// TIA Portal V20 export
// export: Created 2026-10-19T18:44:59.9625904Z, ExportSetting None, DisplayName Totally Integrated Automation Portal, DisplayVersion V20 Update 6, DisplayName TIA Portal Openness, DisplayVersion V20 Update 6, DisplayName TIA Portal Version Control Interface, DisplayVersion V20 Update 6, DisplayName SINAMICS Startdrive Advanced, DisplayVersion V20 SP1, DisplayName SINAMICS Startdrive G130, G150, S120, S150, SINAMICS MV, G220, S200, S210, DisplayVersion V20 SP1, DisplayName SINAMICS Startdrive G110M, G120, G120C, G120D, G120P, G115D, DisplayVersion V20 SP1, DisplayName STEP 7 Professional, DisplayVersion V20 Update 6, DisplayName STEP 7 Safety, DisplayVersion V20 Update 2, DisplayName WinCC Basic/Comfort/Advanced, DisplayVersion V20 Update 6, DisplayName WinCC Unified, DisplayVersion V20 Update 6
VAR_GLOBAL   // PLC tag table "Default tag table"
   System_Byte AT %MB1159 : Byte;
   FirstScan AT %M1159.0 : Bool;
   DiagStatusUpdate AT %M1159.1 : Bool;
   AlwaysTRUE AT %M1159.2 : Bool;
   AlwaysFALSE AT %M1159.3 : Bool;
   Clock_Byte AT %MB1160 : Byte;
   Clock_10Hz AT %M1160.0 : Bool;
   Clock_5Hz AT %M1160.1 : Bool;
   "Clock_2.5Hz" AT %M1160.2 : Bool;
   Clock_2Hz AT %M1160.3 : Bool;
   "Clock_1.25Hz" AT %M1160.4 : Bool;
   Clock_1Hz AT %M1160.5 : Bool;
   "Clock_0.625Hz" AT %M1160.6 : Bool;
   "Clock_0.5Hz" AT %M1160.7 : Bool;
   Tag_1 AT %M2000.0 : Bool;
   Tag_2 AT %M2000.1 : Bool;
   Tag_3 AT %M2000.2 : Bool;
   Reintegration AT %M2000.3 : Bool;
   Error_Word_1 AT %MW2001 : Word;
   "Auto_Stop_Lector(1)" AT %M20.6 : Bool;
   "Auto_Stop_Lector(2)" AT %M20.7 : Bool;
   "Auto_Start_Lector(1)" AT %M19.6 : Bool;
   "Auto_Start_Lector(2)" AT %M20.2 : Bool;
   Force_System_1 AT %M25.5 : Bool;
   VTD_System_Selected_HMI AT %MW1234 : UInt;
   Initialization AT %M19.4 : Bool;
   Save_Settings AT %M0.1 : Bool;
   "LE_Bypass(1)" AT %M704.1 : Bool;
   "LE_Bypass(2)" AT %M704.2 : Bool;
   Reset_Comissioning AT %M70.0 : Bool;
   System_2_Busy AT %M39.6 : Bool;
   System_1_Busy AT %M19.5 : Bool;
   L3_OK AT %M39.4 : Bool;
   L4_OK AT %M39.0 : Bool;
   L5_OK AT %M39.1 : Bool;
   L1_OK AT %M26.6 : Bool;
   L2_OK AT %M26.7 : Bool;
   L6_OK AT %M39.2 : Bool;
   L1_Estop AT %M61.6 : Bool;
   L6_Estop AT %M70.6 : Bool;
   L2_Estop AT %M61.7 : Bool;
   L5_Estop AT %M70.4 : Bool;
   L4_Estop AT %M70.3 : Bool;
   L3_Estop AT %M70.2 : Bool;
   LGX_Secure_Access_2 AT %M71.5 : Bool;
   LGX_Secure_Access_1 AT %M71.4 : Bool;
   LGX_ReadyToReceive_2 AT %M71.2 : Bool;
   LGX_ReadyToReceive_1 AT %M61.5 : Bool;
   Dbug AT %M71.7 : Bool;
   OrderNo AT %MW158 : Int;
   "Clear_OT_Buffers(1)" AT %M154.6 : Bool;
   "Clear_OT_Buffers(2)" AT %M154.7 : Bool;
   "Clear_OT_VTD(1)" AT %M154.4 : Bool;
   "Clear_OT_VTD(2)" AT %M154.5 : Bool;
END_VAR
